// TIA Portal V19 export
// export: Created 2026-01-15T10:00:00.0000000Z, ExportSetting WithReadOnly
FUNCTION "FC_ExampleScale" : Void   // FC20, STL
// stored: IsKnowHowProtected false
   VAR_INPUT
      In : Int;
   END_VAR
   VAR_OUTPUT
      Out : Int;
   END_VAR
BEGIN

NETWORK
TITLE = 
      L     #In;
      L     10;
      *I;
      T     #Out;

//scaled by ten
END_FUNCTION
